// TIA Portal V20 export
// export: Created 2026-10-19T18:45:18.6122602Z, ExportSetting None, DisplayName Totally Integrated Automation Portal, DisplayVersion V20 Update 6, DisplayName TIA Portal Openness, DisplayVersion V20 Update 6, DisplayName TIA Portal Version Control Interface, DisplayVersion V20 Update 6, DisplayName SINAMICS Startdrive Advanced, DisplayVersion V20 SP1, DisplayName SINAMICS Startdrive G130, G150, S120, S150, SINAMICS MV, G220, S200, S210, DisplayVersion V20 SP1, DisplayName SINAMICS Startdrive G110M, G120, G120C, G120D, G120P, G115D, DisplayVersion V20 SP1, DisplayName STEP 7 Professional, DisplayVersion V20 Update 6, DisplayName STEP 7 Safety, DisplayVersion V20 Update 2, DisplayName WinCC Basic/Comfort/Advanced, DisplayVersion V20 Update 6, DisplayName WinCC Unified, DisplayVersion V20 Update 6
VAR_GLOBAL   // PLC tag table "IO_Remote_Panel_1"
   "RESET LAMP(1)" AT %Q0.0 : Bool;   // TESTED
   "VTD1 UPPER ULTIMATE CREEP" AT %I1.1 : Bool;
   "Chain Slack 4 - CH2(1)" AT %I321.7 : Bool;
   "KEY REMOTE/LOCAL L2 - CH1(1)" AT %I338.7 : Bool;
   "STO VTD - CH1(1)" AT %Q370.2 : Bool;
   "VTD1 LOWER LIMIT" AT %I1.2 : Bool;
   "KEY REMOTE/LOCAL L5 - CH1(1)" AT %I347.5 : Bool;
   "VTD1 UPPER ULTIMATE SLOWDOWN" AT %I1.0 : Bool;
   "LIGHT GUARDS 2 - CH2(1)" AT %I330.2 : Bool;
   "SAFETY_GATE_1_CH1(1)" AT %I338.0 : Bool;
   "KEY REMOTE/LOCAL L3 - CH2(1)" AT %I348.1 : Bool;
   "E-STOP L1 - CH2(1)" AT %I339.4 : Bool;
   "KEY REMOTE/LOCAL L4 - CH2(1)" AT %I348.3 : Bool;
   "Chain Slack 3 - CH2(1)" AT %I321.6 : Bool;
   "C1101, C1102, C1103, C1104 CIRCUIT BREAKER" AT %I0.1 : Bool;
   "Chain Slack 2 - CH2(1)" AT %I321.5 : Bool;
   "SAFETY_GATE_4_CH2(1)" AT %I339.3 : Bool;
   "E-STOP L2 - CH1(1)" AT %I338.6 : Bool;
   "E-STOP L1 - CH1(1)" AT %I338.4 : Bool;
   "KEY REMOTE/LOCAL L5 - CH2(1)" AT %I348.5 : Bool;
   "VTD1 PUSH TO EXIT VTD ZONE" AT %I1.6 : Bool;
   "KEY REMOTE/LOCAL L1 - CH1(1)" AT %I338.5 : Bool;
   "SAFETY_GATE_4_CH1(1)" AT %I338.3 : Bool;
   "Chain Slack 1 - CH1(1)" AT %I320.4 : Bool;
   "CABINET 24V PSU CIRCUIT BREAKER FEEDBACK_1(1)" AT %I0.6 : Bool;
   "E-STOP L3 - CH1(1)" AT %I347.0 : Bool;
   "KEY REMOTE/LOCAL L2 - CH2(1)" AT %I339.7 : Bool;
   "E-STOP (CABINET) - CH1(1)" AT %I320.0 : Bool;
   "E-STOP L5 - CH1(1)" AT %I347.4 : Bool;
   "LIGHT GUARD 1 - CH1(1)" AT %I329.1 : Bool;
   "VTD1 LOWER ULTIMATE SLOWDOWN" AT %I1.4 : Bool;
   "LIGHT GUARDS 1 - CH2(1)" AT %I330.1 : Bool;
   "E-STOP L3 - CH2(1)" AT %I348.0 : Bool;
   "E-STOP (CABINET) - CH2(1)" AT %I321.0 : Bool;
   "KEY REMOTE/LOCAL L4 - CH1(1)" AT %I347.3 : Bool;
   "VTD1 PUSH TO ENTER VTD ZONE" AT %I1.5 : Bool;
   "C1109, C1110, C1111 CVTD CIRCUIT BREAKER" AT %I0.3 : Bool;
   "BRAKE SUPPLY SAFETY CONTACTOR 1(1)" AT %Q370.0 : Bool;
   "SAFETY_GATE_1_CH2(1)" AT %I339.0 : Bool;
   "KEY REMOTE/LOCAL L3 - CH1(1)" AT %I347.1 : Bool;
   "CABINET COOLING FAN CIRCUIT BREAKER FEEDBACK(1)" AT %I0.4 : Bool;
   "E-STOP L6 - CH2(1)" AT %I348.6 : Bool;
   "Chain Slack 1 - CH2(1)" AT %I321.4 : Bool;
   "E-STOP L4 - CH2(1)" AT %I348.2 : Bool;
   "RESET (CABINET)(1)" AT %I320.1 : Bool;
   "SAFETY_GATE_2_CH1(1)" AT %I338.1 : Bool;
   "E-STOP L4 - CH1(1)" AT %I347.2 : Bool;
   "KEY REMOTE/LOCAL L6 - CH2(1)" AT %I348.7 : Bool;
   "STO VTD - CH2(1)" AT %Q370.3 : Bool;
   "CABINET 24V PSU CIRCUIT BREAKER FEEDBACK(1)" AT %I0.5 : Bool;
   "SAFETY_GATE_3_CH2(1)" AT %I339.2 : Bool;
   "SAFETY_GATE_3_CH1(1)" AT %I338.2 : Bool;
   "E-STOP L2 - CH2(1)" AT %I339.6 : Bool;
   "E-STOP L5 - CH2(1)" AT %I348.4 : Bool;
   "Chain Slack 4 - CH1(1)" AT %I320.7 : Bool;
   "VTU HOIST BRAKE SAFETY ENABLE EDM FEEDBACK(1)" AT %I329.0 : Bool;
   "E-STOP L6 - CH1(1)" AT %I347.6 : Bool;
   "SAFETY_GATE_2_CH2(1)" AT %I339.1 : Bool;
   "KEY REMOTE/LOCAL L1 - CH2(1)" AT %I339.5 : Bool;
   "VTD1 UPPER LIMIT" AT %I1.3 : Bool;
   "Chain Slack 3 - CH1(1)" AT %I320.6 : Bool;
   "BRAKE SUPPLY SAFETY CONTACTOR 2(1)" AT %Q370.1 : Bool;
   "KEY REMOTE/LOCAL L6 - CH1(1)" AT %I347.7 : Bool;
   "LIGHT GUARD 2 - CH1(1)" AT %I329.2 : Bool;
   "C1112 VTD CIRCUIT BREAKER" AT %I0.0 : Bool;
   "Chain Slack 2 - CH1(1)" AT %I320.5 : Bool;
   "C1105, C1106, C1107, C1108 CIRCUIT BREAKER" AT %I0.2 : Bool;
   "STACK LIGHTS GREEN(1)" AT %Q0.3 : Bool;
   "STACK LIGHTS RED(1)" AT %Q0.1 : Bool;
   "STACK LIGHTS ORANGE(1)" AT %Q0.2 : Bool;
END_VAR
